LAYER Default
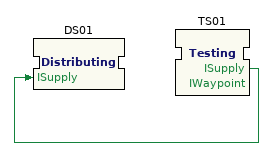
  FBS
    DS01 : Distributing;
    TS01 : Testing;
  END_FBS
  ADAPTER_CONNECTIONS
    TS01.ISupply TO DS01.ISupply;
  END_CONNECTIONS
END_LAYER
